(* PLC project forms.project, CODESYS CODESYS V3.5 SP17 Patch 3 *)
(* stored: creationDateTime 2026-10-20T03:44:11.2858434, modificationDateTime 1601-01-01T03:00:00 *)

{attribute 'qualified_only'}
VAR_GLOBAL  (* GVL_Probe *)
  xFlag : BOOL;
  iCount : INT := 5;
  rTotal : REAL;
  diHours : DINT;
END_VAR
